FUNCTION_BLOCK E_MERGE_5 (* Extracted Composite Function Block Type *)
  (* Standard: 61499-2 *)
  (* Version 10/20/2026, macie *)
  PACKAGE Main;
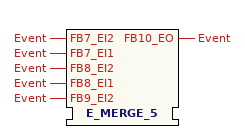
  EVENT_INPUT
    FB7_EI2; (* Second input event *)
    FB7_EI1; (* First input event *)
    FB8_EI2; (* Second input event *)
    FB8_EI1; (* First input event *)
    FB9_EI2; (* Second input event *)
  END_EVENT
  EVENT_OUTPUT
    FB10_EO; (* Output Event *)
  END_EVENT
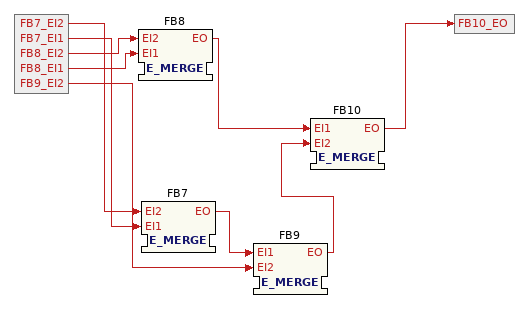
  FBS
    FB7 : E_MERGE;
    FB8 : E_MERGE;
    FB9 : E_MERGE;
    FB10 : E_MERGE;
  END_FBS
  EVENT_CONNECTIONS
    FB7.EO TO FB9.EI1;
    FB8.EO TO FB10.EI1;
    FB9.EO TO FB10.EI2;
    FB7_EI2 TO FB7.EI2;
    FB7_EI1 TO FB7.EI1;
    FB8_EI2 TO FB8.EI2;
    FB8_EI1 TO FB8.EI1;
    FB9_EI2 TO FB9.EI2;
    FB10.EO TO FB10_EO;
  END_CONNECTIONS
END_FUNCTION_BLOCK
